// TIA Portal V20 export
// export: Created 2026-10-20T12:46:36.0742882Z, ExportSetting WithDefaults, DisplayName Totally Integrated Automation Portal, DisplayVersion V20 Update 6, DisplayName TIA Portal Openness, DisplayVersion V20 Update 6, DisplayName TIA Portal Version Control Interface, DisplayVersion V20 Update 6, DisplayName SINAMICS Startdrive Advanced, DisplayVersion V20 SP1, DisplayName SINAMICS Startdrive G130, G150, S120, S150, SINAMICS MV, G220, S200, S210, DisplayVersion V20 SP1, DisplayName SINAMICS Startdrive G110M, G120, G120C, G120D, G120P, G115D, DisplayVersion V20 SP1, DisplayName STEP 7 Professional, DisplayVersion V20 Update 6, DisplayName STEP 7 Safety, DisplayVersion V20 Update 2, DisplayName WinCC Basic/Comfort/Advanced, DisplayVersion V20 Update 6, DisplayName WinCC Unified, DisplayVersion V20 Update 6
DATA_BLOCK "MQTT_Handler_FB_DB"   // DB44
VERSION : 0.1
// stored: AutoNumber true, DBAccessibleFromOPCUA true, InstanceOfName MQTT_Handler_FB, InstanceOfType FB
"MQTT_Handler_FB"
   // VAR_INPUT
   //    Enable : Bool;
   // END_VAR
   // VAR_IN_OUT
   //    LMQTT_DB : "LMQTT_DB_UDT";
   // END_VAR
   // VAR
   //    MQTT_Setup : Bool;
   //    MQTT_Topic : WString;
   //    Publish_Msg_Payload : Array[1..128] of Byte;
   //    Received_Topic : WString;
   //    Received_Msg_Payload : Array[0..1024] of Byte;
   //    i : UInt;
   //    j : UInt;
   //    Subscribe : Bool;
   //    Unsubscribe : Bool;
   //    Received_Msg_Status : USInt;
   //    Received_Msg_Length : UDInt;
   //    Busy : Bool;
   //    Valid : Bool;
   //    Done : Bool;
   //    Error : Bool;
   //    Status : Word;
   //    Diagnostics { S7_SetPoint := 'True'} : "typeDiagnostics";
   //    JSON_Tree : Array[1..18] of "LStream_typeElement";
   //    Shuttle_No : UInt;
   //    sSubTopic : Array[1..24] of String;
   //    bSubscribed : Bool;
   //    SubscribeState : Int;
   //    SubscribeIndex : Int;
   //    SubscribeCount : UInt;
   //    SubscribeTopicList : Array[1..30] of String;
   //    sPayloadRcv : String;
   //    sPayloadRcv_1 : String;
   //    sPayloadRcv_2 : String;
   //    sPayloadRcv_3 : String;
   //    sPayloadRcv_4 : String;
   //    sPayloadRcv_5 : String;
   //    MQTT_AutoReset : UInt;
   //    Enable_AutoReset : Bool;
   //    T_AutoReset { S7_SetPoint := 'True'} : TON_TIME;
   // END_VAR
BEGIN
END_DATA_BLOCK
